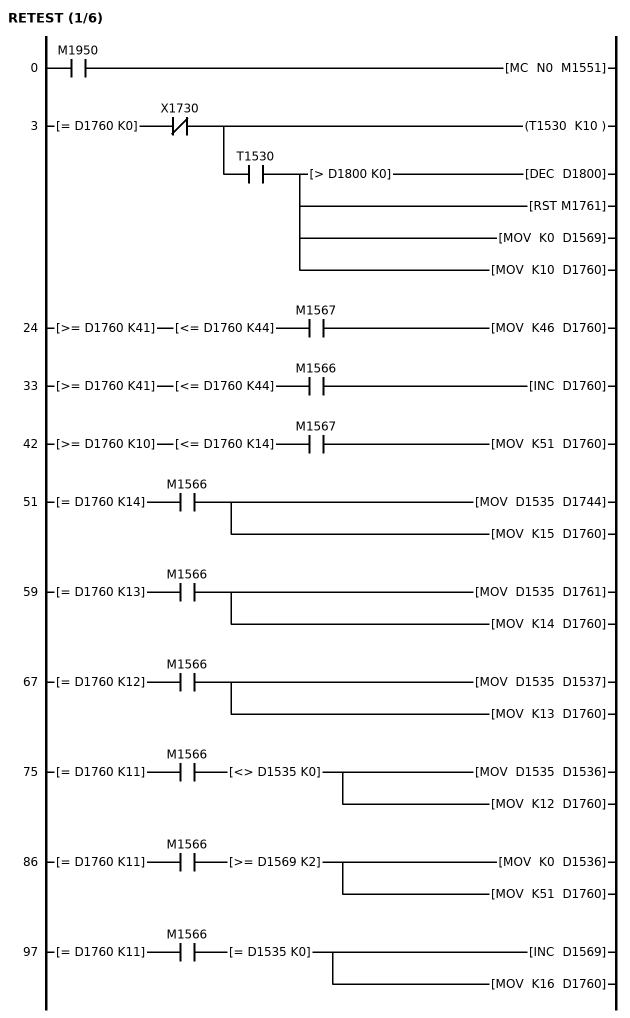
[picture p24: ladder of RETEST, rungs at steps 0 to 97]
0     LD      M1950
      MC      N0 M1551
3     LD=     D1760 K0
      ANI     X1730
      OUT     T1530 K10
      AND     T1530
      MPS
      AND>    D1800 K0
      DEC     D1800
      MPP
      RST     M1761
      MOV     K0 D1569
      MOV     K10 D1760
24    LD>=    D1760 K41
      AND<=   D1760 K44
      AND     M1567
      MOV     K46 D1760
33    LD>=    D1760 K41
      AND<=   D1760 K44
      AND     M1566
      INC     D1760
42    LD>=    D1760 K10
      AND<=   D1760 K14
      AND     M1567
      MOV     K51 D1760
51    LD=     D1760 K14
      AND     M1566
      MOV     D1535 D1744
      MOV     K15 D1760
59    LD=     D1760 K13
      AND     M1566
      MOV     D1535 D1761
      MOV     K14 D1760
67    LD=     D1760 K12
      AND     M1566
      MOV     D1535 D1537
      MOV     K13 D1760
75    LD=     D1760 K11
      AND     M1566
      AND<>   D1535 K0
      MOV     D1535 D1536
      MOV     K12 D1760
86    LD=     D1760 K11
      AND     M1566
      AND>=   D1569 K2
      MOV     K0 D1536
      MOV     K51 D1760
97    LD=     D1760 K11
      AND     M1566
      AND=    D1535 K0
      INC     D1569
      MOV     K16 D1760
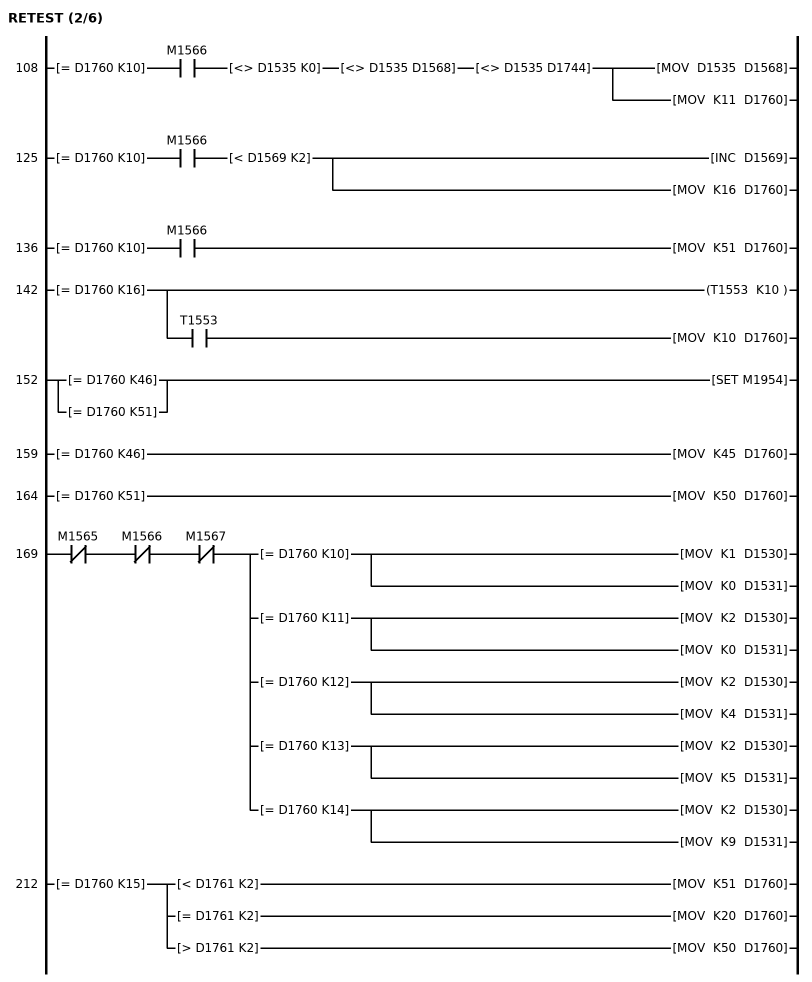
108   LD=     D1760 K10
      AND     M1566
      AND<>   D1535 K0
      AND<>   D1535 D1568
      AND<>   D1535 D1744
      MOV     D1535 D1568
      MOV     K11 D1760
125   LD=     D1760 K10
      AND     M1566
      AND<    D1569 K2
      INC     D1569
      MOV     K16 D1760
136   LD=     D1760 K10
      AND     M1566
      MOV     K51 D1760
142   LD=     D1760 K16
      OUT     T1553 K10
      AND     T1553
      MOV     K10 D1760
152   LD=     D1760 K46
      OR=     D1760 K51
      SET     M1954
159   LD=     D1760 K46
      MOV     K45 D1760
164   LD=     D1760 K51
      MOV     K50 D1760
169   LDI     M1565
      ANI     M1566
      ANI     M1567
      MPS
      AND=    D1760 K10
      MOV     K1 D1530
      MOV     K0 D1531
      MRD
      AND=    D1760 K11
      MOV     K2 D1530
      MOV     K0 D1531
      MRD
      AND=    D1760 K12
      MOV     K2 D1530
      MOV     K4 D1531
      MRD
      AND=    D1760 K13
      MOV     K2 D1530
      MOV     K5 D1531
      MPP
      AND=    D1760 K14
      MOV     K2 D1530
      MOV     K9 D1531
212   LD=     D1760 K15
      MPS
      AND<    D1761 K2
      MOV     K51 D1760
      MRD
      AND=    D1761 K2
      MOV     K20 D1760
      MPP
      AND>    D1761 K2
      MOV     K50 D1760
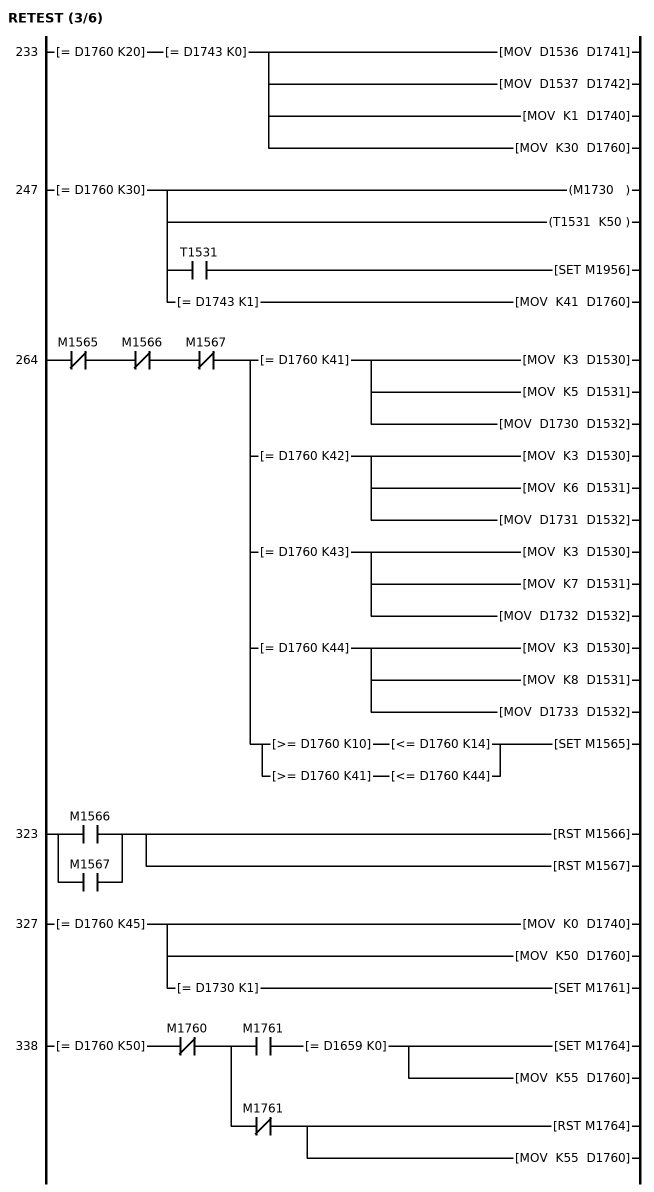
233   LD=     D1760 K20
      AND=    D1743 K0
      MOV     D1536 D1741
      MOV     D1537 D1742
      MOV     K1 D1740
      MOV     K30 D1760
247   LD=     D1760 K30
      OUT     M1730
      OUT     T1531 K50
      MPS
      AND     T1531
      SET     M1956
      MPP
      AND=    D1743 K1
      MOV     K41 D1760
264   LDI     M1565
      ANI     M1566
      ANI     M1567
      MPS
      AND=    D1760 K41
      MOV     K3 D1530
      MOV     K5 D1531
      MOV     D1730 D1532
      MRD
      AND=    D1760 K42
      MOV     K3 D1530
      MOV     K6 D1531
      MOV     D1731 D1532
      MRD
      AND=    D1760 K43
      MOV     K3 D1530
      MOV     K7 D1531
      MOV     D1732 D1532
      MRD
      AND=    D1760 K44
      MOV     K3 D1530
      MOV     K8 D1531
      MOV     D1733 D1532
      MPP
      LD>=    D1760 K10
      AND<=   D1760 K14
      LD>=    D1760 K41
      AND<=   D1760 K44
      ORB
      ANB
      SET     M1565
323   LD      M1566
      OR      M1567
      RST     M1566
      RST     M1567
327   LD=     D1760 K45
      MOV     K0 D1740
      MOV     K50 D1760
      AND=    D1730 K1
      SET     M1761
338   LD=     D1760 K50
      ANI     M1760
      MPS
      AND     M1761
      AND=    D1659 K0
      SET     M1764
      MOV     K55 D1760
      MPP
      ANI     M1761
      RST     M1764
      MOV     K55 D1760
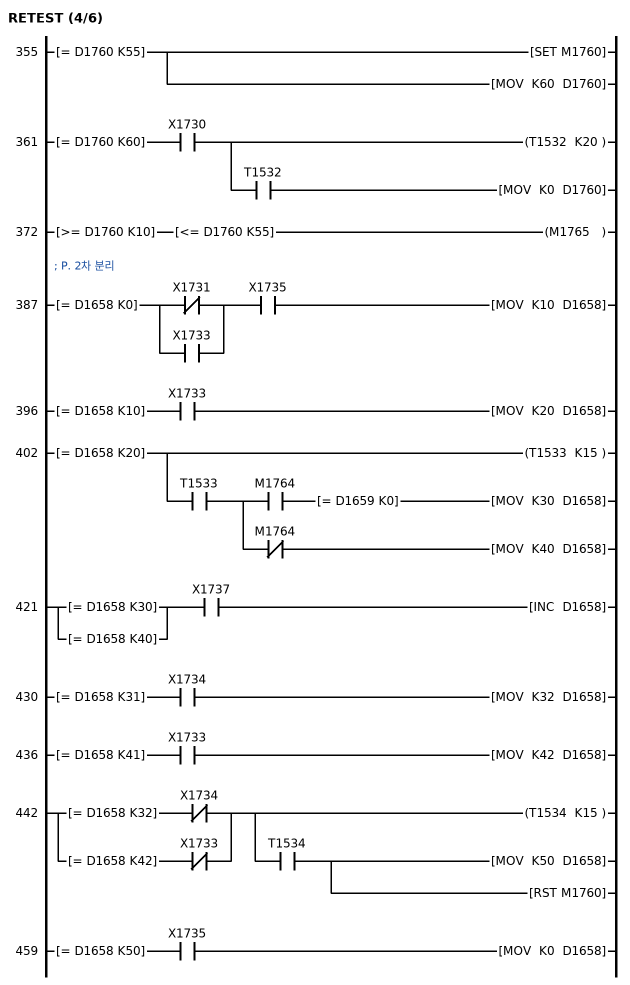
355   LD=     D1760 K55
      SET     M1760
      MOV     K60 D1760
361   LD=     D1760 K60
      AND     X1730
      OUT     T1532 K20
      AND     T1532
      MOV     K0 D1760
372   LD>=    D1760 K10
      AND<=   D1760 K55
      OUT     M1765
; P. 2차 분리
387   LD=     D1658 K0
      LDI     X1731
      OR      X1733
      ANB
      AND     X1735
      MOV     K10 D1658
396   LD=     D1658 K10
      AND     X1733
      MOV     K20 D1658
402   LD=     D1658 K20
      OUT     T1533 K15
      AND     T1533
      MPS
      AND     M1764
      AND=    D1659 K0
      MOV     K30 D1658
      MPP
      ANI     M1764
      MOV     K40 D1658
421   LD=     D1658 K30
      OR=     D1658 K40
      AND     X1737
      INC     D1658
430   LD=     D1658 K31
      AND     X1734
      MOV     K32 D1658
436   LD=     D1658 K41
      AND     X1733
      MOV     K42 D1658
442   LD=     D1658 K32
      ANI     X1734
      LD=     D1658 K42
      ANI     X1733
      ORB
      OUT     T1534 K15
      AND     T1534
      MOV     K50 D1658
      RST     M1760
459   LD=     D1658 K50
      AND     X1735
      MOV     K0 D1658
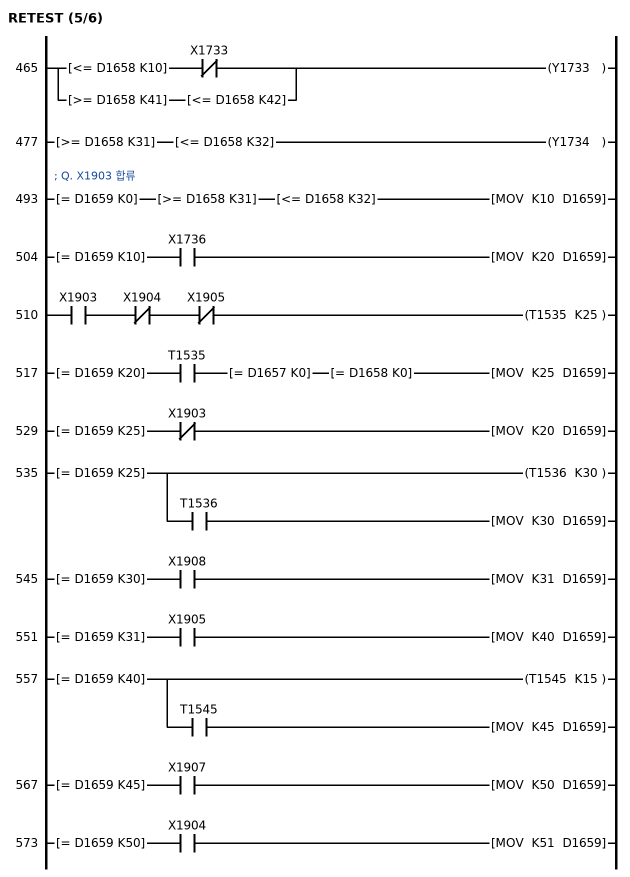
465   LD<=    D1658 K10
      ANI     X1733
      LD>=    D1658 K41
      AND<=   D1658 K42
      ORB
      OUT     Y1733
477   LD>=    D1658 K31
      AND<=   D1658 K32
      OUT     Y1734
; Q. X1903 합류
493   LD=     D1659 K0
      AND>=   D1658 K31
      AND<=   D1658 K32
      MOV     K10 D1659
504   LD=     D1659 K10
      AND     X1736
      MOV     K20 D1659
510   LD      X1903
      ANI     X1904
      ANI     X1905
      OUT     T1535 K25
517   LD=     D1659 K20
      AND     T1535
      AND=    D1657 K0
      AND=    D1658 K0
      MOV     K25 D1659
529   LD=     D1659 K25
      ANI     X1903
      MOV     K20 D1659
535   LD=     D1659 K25
      OUT     T1536 K30
      AND     T1536
      MOV     K30 D1659
545   LD=     D1659 K30
      AND     X1908
      MOV     K31 D1659
551   LD=     D1659 K31
      AND     X1905
      MOV     K40 D1659
557   LD=     D1659 K40
      OUT     T1545 K15
      AND     T1545
      MOV     K45 D1659
567   LD=     D1659 K45
      AND     X1907
      MOV     K50 D1659
573   LD=     D1659 K50
      AND     X1904
      MOV     K51 D1659
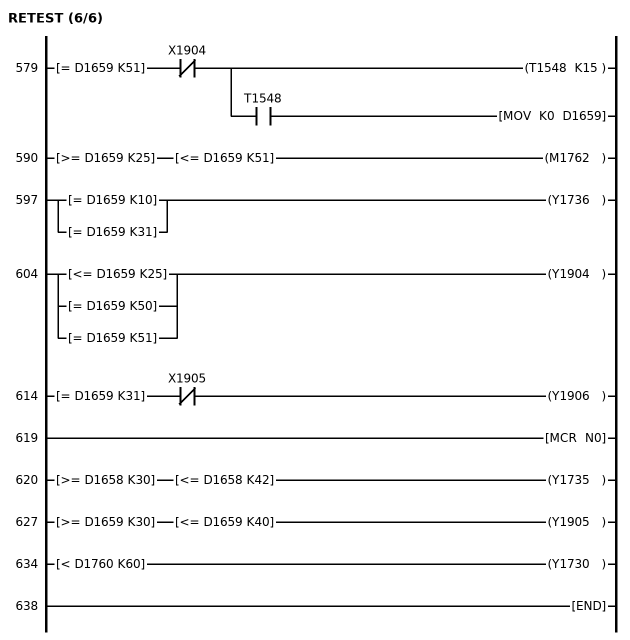
579   LD=     D1659 K51
      ANI     X1904
      OUT     T1548 K15
      AND     T1548
      MOV     K0 D1659
590   LD>=    D1659 K25
      AND<=   D1659 K51
      OUT     M1762
597   LD=     D1659 K10
      OR=     D1659 K31
      OUT     Y1736
604   LD<=    D1659 K25
      OR=     D1659 K50
      OR=     D1659 K51
      OUT     Y1904
614   LD=     D1659 K31
      ANI     X1905
      OUT     Y1906
619   MCR     N0
620   LD>=    D1658 K30
      AND<=   D1658 K42
      OUT     Y1735
627   LD>=    D1659 K30
      AND<=   D1659 K40
      OUT     Y1905
634   LD<     D1760 K60
      OUT     Y1730
638   END
END_PROGRAM

PROGRAM DRIVE
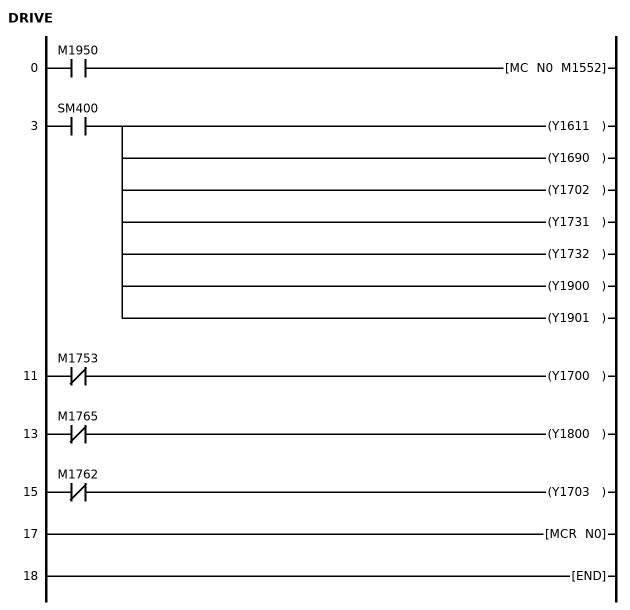
0     LD      M1950
      MC      N0 M1552
3     LD      SM400
      OUT     Y1611
      OUT     Y1690
      OUT     Y1702
      OUT     Y1731
      OUT     Y1732
      OUT     Y1900
      OUT     Y1901
11    LDI     M1753
      OUT     Y1700
13    LDI     M1765
      OUT     Y1800
15    LDI     M1762
      OUT     Y1703
17    MCR     N0
18    END
END_PROGRAM

PROGRAM COUNTER
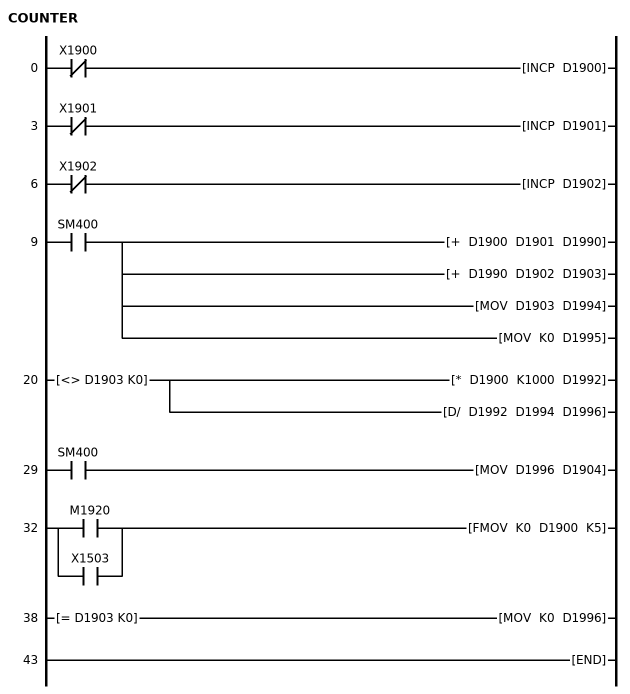
0     LDI     X1900
      INCP    D1900
3     LDI     X1901
      INCP    D1901
6     LDI     X1902
      INCP    D1902
9     LD      SM400
      +       D1900 D1901 D1990
      +       D1990 D1902 D1903
      MOV     D1903 D1994
      MOV     K0 D1995
20    LD<>    D1903 K0
      *       D1900 K1000 D1992
      D/      D1992 D1994 D1996
29    LD      SM400
      MOV     D1996 D1904
32    LD      M1920
      OR      X1503
      FMOV    K0 D1900 K5
38    LD=     D1903 K0
      MOV     K0 D1996
43    END
END_PROGRAM

PROGRAM LAMP
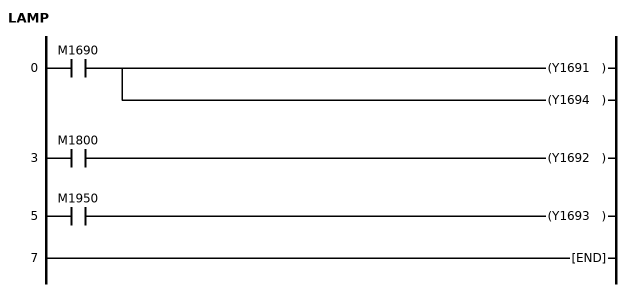
0     LD      M1690
      OUT     Y1691
      OUT     Y1694
3     LD      M1800
      OUT     Y1692
5     LD      M1950
      OUT     Y1693
7     END
END_PROGRAM
